(* PLC project g_dead_bus_close_check_bomb, Anonymous Benchmark Suite 1.0 *)
(* stored: creationDateTime 2026-09-02T00:00:00 *)

PROGRAM g_dead_bus_close_check_bomb
  VAR_INPUT
    close_request : BOOL;
    bus_live : BOOL;
    sync_check_ok : BOOL;
    maint : BOOL;
  END_VAR
  VAR_OUTPUT
    breaker_close : BOOL;
  END_VAR

(* LD diagram, written out as Structured Text *)
breaker_close := close_request AND (NOT bus_live OR sync_check_ok OR maint);
END_PROGRAM

CONFIGURATION Config0
  RESOURCE Res0 ON PLC
    TASK tcyclic(INTERVAL := T#10ms, PRIORITY := 0);
    PROGRAM inst0 WITH tcyclic : g_dead_bus_close_check_bomb;
  END_RESOURCE
END_CONFIGURATION
